SUBAPPLICATION Uebung_OPC_L11_AX (* Wie Training_11, lokal: SoftKeys F1/F2 statt Tastern, erreichter Zustand lokal zurueck auf den SoftKey-Hintergrund *)
  (* Standard: 61499-2; Description: Copyright (c) 2026 Meisterschulen am Ostbahnhof This program and the accompanying materials are made available under the terms of the Eclipse Public License 2.0 which is available at https://www.eclipse.org/legal/epl-2.0/ SPDX-License-Identifier: EPL-2.0 *)
  (* Version 1.0, 2026-10-18, Franz Höpfinger, Meisterschulen am Ostbahnhof, Aus SubApp_PC_A + SubApp_PC_B von test_VV zusammengefuehrt, lokale Varianten der Bausteine *)
  PACKAGE Meins::OPC_UA_Lokal;
  IMPORT Uebungen::const::UT::DefaultPool::SoftKey_F1;
  IMPORT Uebungen::const::UT::DefaultPool::SoftKey_F2;
  IMPORT Meins::OPC_UA_Lokal::const::OpcUaLokal::SW1_UP_WRITE;
  IMPORT Meins::OPC_UA_Lokal::const::OpcUaLokal::SW1_DOWN_WRITE;
  IMPORT Meins::OPC_UA_Lokal::const::OpcUaLokal::SW1_UP_STATE_READ;
  IMPORT Meins::OPC_UA_Lokal::const::OpcUaLokal::SW1_DOWN_STATE_READ;
  IMPORT Meins::OPC_UA_Lokal::const::OpcUaLokal::SW1_UP_READ;
  IMPORT Meins::OPC_UA_Lokal::const::OpcUaLokal::SW1_DOWN_READ;
  IMPORT Meins::OPC_UA_Lokal::const::OpcUaLokal::SW1_UP_STATE_WRITE;
  IMPORT Meins::OPC_UA_Lokal::const::OpcUaLokal::SW1_DOWN_STATE_WRITE;
  IMPORT logiBUS::io::DQ::logiBUS_DO::Output_Q7;
  IMPORT logiBUS::io::DQ::logiBUS_DO::Output_Q8;
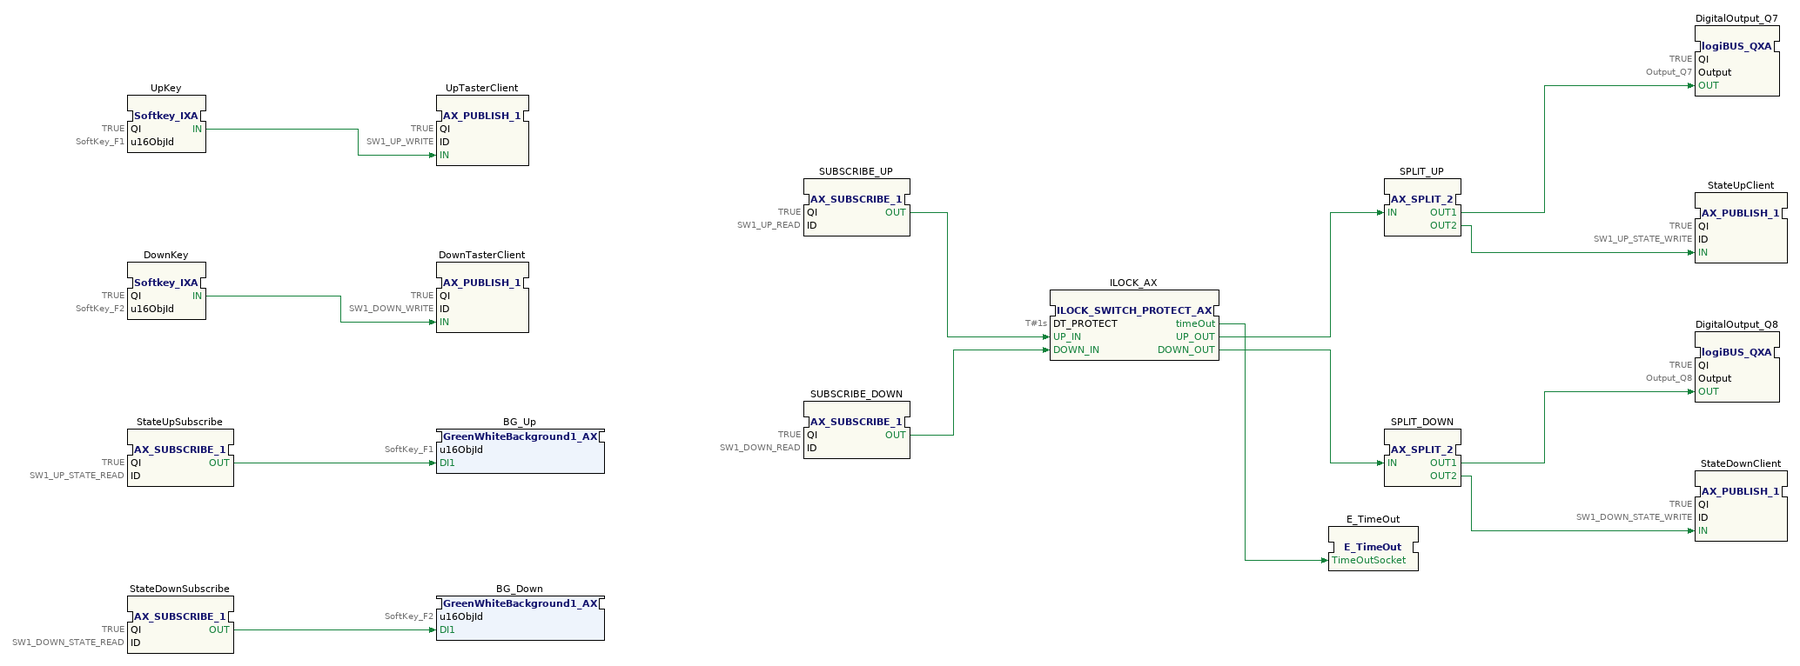
  FBS
    UpKey : isobus::UT::io::Softkey::Softkey_IXA(QI := TRUE, u16ObjId := SoftKey_F1);
    DownKey : isobus::UT::io::Softkey::Softkey_IXA(QI := TRUE, u16ObjId := SoftKey_F2);
    UpTasterClient : adapter::net::AX_PUBLISH_1(QI := TRUE, ID := SW1_UP_WRITE);
    DownTasterClient : adapter::net::AX_PUBLISH_1(QI := TRUE, ID := SW1_DOWN_WRITE);
    StateUpSubscribe : adapter::net::AX_SUBSCRIBE_1(QI := TRUE, ID := SW1_UP_STATE_READ);
    StateDownSubscribe : adapter::net::AX_SUBSCRIBE_1(QI := TRUE, ID := SW1_DOWN_STATE_READ);
    SUBSCRIBE_UP : adapter::net::AX_SUBSCRIBE_1(QI := TRUE, ID := SW1_UP_READ);
    SUBSCRIBE_DOWN : adapter::net::AX_SUBSCRIBE_1(QI := TRUE, ID := SW1_DOWN_READ);
    ILOCK_AX : logiBUS::signalprocessing::interlock::ILOCK_SWITCH_PROTECT_AX(DT_PROTECT := T#1s);
    E_TimeOut : iec61499::events::E_TimeOut;
    SPLIT_UP : adapter::events::unidirectional::AX_SPLIT_2;
    SPLIT_DOWN : adapter::events::unidirectional::AX_SPLIT_2;
    DigitalOutput_Q7 : logiBUS::io::DQ::logiBUS_QXA(QI := TRUE, Output := Output_Q7);
    DigitalOutput_Q8 : logiBUS::io::DQ::logiBUS_QXA(QI := TRUE, Output := Output_Q8);
    StateUpClient : adapter::net::AX_PUBLISH_1(QI := TRUE, ID := SW1_UP_STATE_WRITE);
    StateDownClient : adapter::net::AX_PUBLISH_1(QI := TRUE, ID := SW1_DOWN_STATE_WRITE);
  END_FBS
  SUBAPPS
    BG_Up : MyLib::sys::GreenWhiteBackground1_AX(u16ObjId := SoftKey_F1);
    BG_Down : MyLib::sys::GreenWhiteBackground1_AX(u16ObjId := SoftKey_F2);
  END_SUBAPPS
  ADAPTER_CONNECTIONS
    UpKey.IN TO UpTasterClient.IN;
    DownKey.IN TO DownTasterClient.IN;
    StateUpSubscribe.OUT TO BG_Up.DI1;
    StateDownSubscribe.OUT TO BG_Down.DI1;
    SUBSCRIBE_UP.OUT TO ILOCK_AX.UP_IN;
    SUBSCRIBE_DOWN.OUT TO ILOCK_AX.DOWN_IN;
    ILOCK_AX.timeOut TO E_TimeOut.TimeOutSocket;
    ILOCK_AX.UP_OUT TO SPLIT_UP.IN;
    SPLIT_UP.OUT1 TO DigitalOutput_Q7.OUT;
    SPLIT_UP.OUT2 TO StateUpClient.IN;
    ILOCK_AX.DOWN_OUT TO SPLIT_DOWN.IN;
    SPLIT_DOWN.OUT1 TO DigitalOutput_Q8.OUT;
    SPLIT_DOWN.OUT2 TO StateDownClient.IN;
  END_CONNECTIONS
END_SUBAPPLICATION
